// Mitsubishi GX Works2 project: W_test   PLC: Q03UDE

PROGRAM MAIN
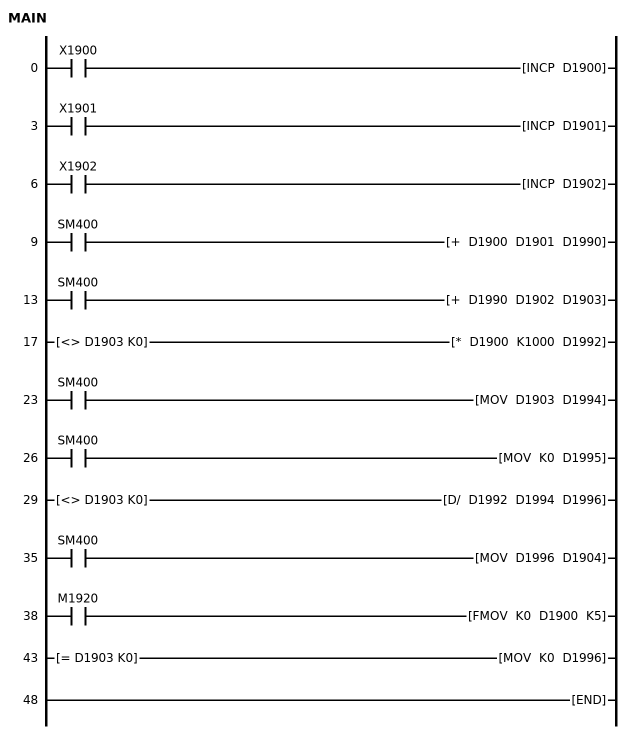
0     LD      X1900
      INCP    D1900
3     LD      X1901
      INCP    D1901
6     LD      X1902
      INCP    D1902
9     LD      SM400
      +       D1900 D1901 D1990
13    LD      SM400
      +       D1990 D1902 D1903
17    LD<>    D1903 K0
      *       D1900 K1000 D1992
23    LD      SM400
      MOV     D1903 D1994
26    LD      SM400
      MOV     K0 D1995
29    LD<>    D1903 K0
      D/      D1992 D1994 D1996
35    LD      SM400
      MOV     D1996 D1904
38    LD      M1920
      FMOV    K0 D1900 K5
43    LD=     D1903 K0
      MOV     K0 D1996
48    END
END_PROGRAM
